(* CODESYS project demo_RECOVERED_2026-10-14T16-49-24.project
   Author: Schneider
   Version: 1.0.0.0

Project tree, tasks and I/O mapping:
  MyController : TM310MM35ECT16U, Schneider Electric, order no. Schneider M310M Target, version 2.0.0.43
    application Application
      libraries: Util, 3.5.19.0 (System); Standard, 3.5.18.0 (System); MC_Basic, 1.10.1.65 (Schneider Electric SA); M310M PLCSystem, * (Schneider Electric)
      task MAST (cyclic, interval T#20ms, priority 15) calls PLC_PRG
      task CommunicationTask (cyclic, interval t#20ms, priority 16) calls nothing
      task MotionTask (cyclic, interval T#4ms, priority 0) calls Motion_PRG, Hidden_PRG
      ImplicitChecks/
        function CheckDivDInt [ST]
        function CheckBounds [ST]
        function CheckLRangeUnsigned [ST]
        function CheckRangeUnsigned [ST]
        function CheckDivReal [ST]
        function CheckDivLReal [ST]
        function CheckRangeSigned [ST]
        function CheckPointer [ST]
        function CheckLRangeSigned [ST]
        function CheckDivLInt [ST]
      program PLC_PRG [ST]
      program Hidden_PRG [ST]
      global variables GVL
      program Motion_PRG [ST]
    Encoders : Encoders, Schneider Electric, version 2.0.0.43
    Cartridge_1 : Cartridge, Schneider Electric, version 2.0.0.43
    IO_Bus : IO bus - TM3, Schneider Electric, version 2.0.0.43
      Module_1 : TM3DI16/G, Schneider Electric, order no. TM3DI16/G, version 1.0.2.2
          input  iwModule_4_IW0 : WORD  // IW0
      Module_2 : TM3DQ16R/G, Schneider Electric, order no. TM3DQ16R/G, version 1.0.2.2
          unmapped channels: QW0
      Module_3 : TM3AI4/G, Schneider Electric, order no. TM3AI4/G, version 1.0.2.2
          settings: KPI Configuration.KPI Configuration = 35; KPI Configuration.KPI Configuration = 160; KPI Configuration.KPI Configuration = 15; KPI Configuration.KPI Configuration = 32; KPI Configuration.KPI Configuration = 78
          input  Application.Motion_PRG.WaterLevel AT %IW3 : INT  // IW0
          input  ibModule_1_IBStatusIW0 : BYTE  // IBStatusIW0
          input  ibModule_1_IBStatusIW1 : BYTE  // IBStatusIW1
          input  ibModule_1_IBStatusIW2 : BYTE  // IBStatusIW2
          input  ibModule_1_IBStatusIW3 : BYTE  // IBStatusIW3
          unmapped channels: %IW4 IW1, %IW5 IW2, IW3
      Module_4 : TM3AQ2/G, Schneider Electric, order no. TM3AQ2/G, version 1.0.2.2
          settings: KPI Configuration.KPI Configuration = 19; KPI Configuration.KPI Configuration = 160; KPI Configuration.KPI Configuration = 15; KPI Configuration.KPI Configuration = 32; KPI Configuration.KPI Configuration = 78
          output qiModule_2_QW1 : INT  // QW1
          input  ibModule_2_IBStatusQW0 : BYTE  // IBStatusQW0
          input  ibModule_2_IBStatusQW1 : BYTE  // IBStatusQW1
          unmapped channels: %QW3 QW0
    EtherCAT_Master_SE : EtherCAT Master SE, Schneider Electric SA, version 4.9.0.3
    Cartridge_2 : Cartridge, Schneider Electric, version 2.0.0.43
    Ethernet_1 : Ethernet Network, Schneider Electric, version 4.3.0.6
        settings: IPAddress = [192,168,0,122]; SubnetMask = [255,255,255,0]; GatewayAddress = [192,168,0,1]; MACAddress = [16#00,16#00,16#00,16#00,16#00,16#00]; IPAddress = [192,168,0,2]; SubnetMask = [255,255,255,0]; GatewayAddress = [0,0,0,0]
      ModbusTCP_Server_Device : ModbusTCP Server Device, Schneider Electric SA, version 4.5.0.1
          input  iwModbusTCP_Server_Device_0 : WORD  // 保持寄存器.保持寄存器
          input  iwModbusTCP_Server_Device_1 : WORD  // 保持寄存器.保持寄存器
          input  iwModbusTCP_Server_Device_2 : WORD  // 保持寄存器.保持寄存器
          input  iwModbusTCP_Server_Device_3 : WORD  // 保持寄存器.保持寄存器
          input  iwModbusTCP_Server_Device_4 : WORD  // 保持寄存器.保持寄存器
          input  iwModbusTCP_Server_Device_5 : WORD  // 保持寄存器.保持寄存器
          input  iwModbusTCP_Server_Device_6 : WORD  // 保持寄存器.保持寄存器
          input  iwModbusTCP_Server_Device_7 : WORD  // 保持寄存器.保持寄存器
          input  iwModbusTCP_Server_Device_8 : WORD  // 保持寄存器.保持寄存器
          input  iwModbusTCP_Server_Device_9 : WORD  // 保持寄存器.保持寄存器
          input  iwModbusTCP_Server_Device_10 : WORD  // 保持寄存器.保持寄存器
          input  iwModbusTCP_Server_Device_11 : WORD  // 保持寄存器.保持寄存器
          input  iwModbusTCP_Server_Device_12 : WORD  // 保持寄存器.保持寄存器
          input  iwModbusTCP_Server_Device_13 : WORD  // 保持寄存器.保持寄存器
          input  iwModbusTCP_Server_Device_14 : WORD  // 保持寄存器.保持寄存器
          input  iwModbusTCP_Server_Device_15 : WORD  // 保持寄存器.保持寄存器
          output qwModbusTCP_Server_Device_0 : WORD  // 输入寄存器.输入寄存器
          output qwModbusTCP_Server_Device_1 : WORD  // 输入寄存器.输入寄存器
          output qwModbusTCP_Server_Device_2 : WORD  // 输入寄存器.输入寄存器
          output qwModbusTCP_Server_Device_3 : WORD  // 输入寄存器.输入寄存器
          output qwModbusTCP_Server_Device_4 : WORD  // 输入寄存器.输入寄存器
          output qwModbusTCP_Server_Device_5 : WORD  // 输入寄存器.输入寄存器
          output qwModbusTCP_Server_Device_6 : WORD  // 输入寄存器.输入寄存器
          output qwModbusTCP_Server_Device_7 : WORD  // 输入寄存器.输入寄存器
          output qwModbusTCP_Server_Device_8 : WORD  // 输入寄存器.输入寄存器
          output qwModbusTCP_Server_Device_9 : WORD  // 输入寄存器.输入寄存器
          output qwModbusTCP_Server_Device_10 : WORD  // 输入寄存器.输入寄存器
          output qwModbusTCP_Server_Device_11 : WORD  // 输入寄存器.输入寄存器
          output qwModbusTCP_Server_Device_12 : WORD  // 输入寄存器.输入寄存器
          output qwModbusTCP_Server_Device_13 : WORD  // 输入寄存器.输入寄存器
          output qwModbusTCP_Server_Device_14 : WORD  // 输入寄存器.输入寄存器
          output qwModbusTCP_Server_Device_15 : WORD  // 输入寄存器.输入寄存器
          unmapped channels: 保持寄存器, 输入寄存器
    Pulse_Generators : Pulse Generators, Schneider Electric, version 2.0.0.43
    Virtual Axis Pool
    COM_1 : Serial COM, Schneider Electric, version 2.0.0.43
    DI : Digital Inputs, Schneider Electric, version 2.0.0.43
        input  iwDI_IW0 : WORD  // IW0
        input  ibDI_IB1 : BYTE  // IB1
    Counters : Counters, Schneider Electric, version 2.0.0.43
    DQ : Digital Outputs, Schneider Electric, version 2.0.0.43
        output qwDQ_QW0 : WORD  // QW0
        output qbDQ_QB1 : BYTE  // QB1
*)

// MyController/Application/GVL
{attribute 'qualified_only'}
VAR_GLOBAL
	rTargetLevel AT %MW0   : REAL := 40.0;    (* 目标水位 %, 占 MW0-1 *)
    rManualValve AT %MW2   : REAL := 0.0;     (* 手动阀开度 %, 占 MW2-3 *)

    (* ===== 状态/报警 (只读供 HMI) ===== *)
	rLevel       AT %MW4   : REAL;     (* 实测水位 %, 占 MW4-5 *)
	rValveCmd    AT %MW6   : REAL;     (* 阀指令 %, 占 MW6-7 *)
END_VAR

// MyController/Application/PLC_PRG
PROGRAM PLC_PRG
VAR
	    (* ===== 周期 ===== *)
    tCycle : TIME := T#100MS;
    rDt    : REAL;                       (* 采样周期, 秒 *)

    (* ===== 物理IO (地址须与 Device IO Mapping 核对) ===== *)
    iLevelRaw AT %IW3    : INT;          (* 水位 4-20mA, 4000..20000 = 0..100% *)
    iValveOut  AT %QW3   : INT;          (* 抽水阀开度 4-20mA, 4000..20000 = 0..100% *)
    bPump      AT %QX4.0 : BOOL;         (* 抽水泵继电器, ON=抽水 *)

    (* ===== HMI / Modbus 设定 (地址可按需调整) ===== *)
    //rTargetLevel AT %MW0   : REAL := 40.0;    (* 目标水位 %, 占 MW0-1 *)
    bAuto        AT %MX102.0 : BOOL := TRUE;    (* 1=自动 0=手动 *)
   // rManualValve AT %MW2   : REAL := 0.0;     (* 手动阀开度 %, 占 MW2-3 *)
    bManualPump  AT %MX106.0 : BOOL := FALSE;   (* 手动泵 ON *)

    (* ===== 状态/报警 (只读供 HMI) ===== *)
	//rLevel       AT %MW4   : REAL;     (* 实测水位 %, 占 MW4-5 *)
	//rValveCmd    AT %MW6   : REAL;     (* 阀指令 %, 占 MW6-7 *)
    bPumpCmd     AT %MX114.0 : BOOL;     (* 泵指令 *)
    bSensorFault AT %MX114.1 : BOOL;     (* 传感器故障 *)
    bAlarm       AT %MX114.2 : BOOL;     (* 总报警 *)

    (* ===== 量程 (INT) ===== *)
    iRawMin : INT := 4000;
    iRawMax : INT := 20000;

    (* ===== PID 内部 ===== *)
    rError, rPrevError, rInt, rDeriv, rPD, rOut : REAL;

    (* ===== PID 参数 (待整定, 见文档) ===== *)
    //rKp : REAL := 3.0;
   // rKi : REAL := 0.1;     (* 1/s, 抵消自然入流静差; 积分对象 Ki 勿过大 *)
   // rKd : REAL := 0.0;
	rKp AT %MW20 : REAL := 3.0;      (* 占 MW20-21, 默认值(上电/未使能时用) *)
    rKi AT %MW22 : REAL := 0.5;      (* 占 MW22-23 *)
    rKd AT %MW24 : REAL := 0.0;      (* 占 MW24-25 *)
    bPidTune : BOOL := FALSE;        (* 1=采用 Modbus 传入的 Kp/Ki/Kd, 0=用上面默认 *)

    (* ===== 联锁阈值 (%, 工程量) ===== *)
    rLvlHH      : REAL := 95.0;   (* 高高: 最大抽水降压 *)
    rLvlLL      : REAL := 5.0;    (* 低低: 停泵防干抽, 靠自流回涨 *)
    rPumpOnThr  : REAL := 3.0;    (* 阀开度>3% 开泵 *)
    rPumpOffThr : REAL := 1.0;    (* 阀开度<1% 关泵(防憋压) *)
	
END_VAR

rDt := TIME_TO_REAL(tCycle) / 1000;   (* 0.1 s *)
(* ===== Modbus 读入: 上位机 -> PLC 设定值 ===== *)
(* REAL 占 2 字, 低字在前(Device_0=低字, 与现有 rLevel 映射顺序一致) *)
%MW0 := iwModbusTCP_Server_Device_0;   (* rTargetLevel 低字 *)
%MW1 := iwModbusTCP_Server_Device_1;   (* rTargetLevel 高字 *)
%MW2 := iwModbusTCP_Server_Device_6;   (* rManualValve 低字 (可选) *)
%MW3 := iwModbusTCP_Server_Device_7;   (* rManualValve 高字 (可选) *)
bAuto       := iwModbusTCP_Server_Device_10.0;   (* 提取 bit0 *)
bManualPump := iwModbusTCP_Server_Device_10.1;   (* 提取 bit1 *)
bPidTune    := iwModbusTCP_Server_Device_10.2;   (* 提取 bit2 *)

(* 仅当使能位置 1 时, 才用 Modbus 传入的 PID 参数覆盖默认值 *)
IF bPidTune THEN
    %MW20 := iwModbusTCP_Server_Device_2;    (* rKp 低字 *)
    %MW21 := iwModbusTCP_Server_Device_3;    (* rKp 高字 *)
    %MW22 := iwModbusTCP_Server_Device_4;    (* rKi 低字 *)
    %MW23 := iwModbusTCP_Server_Device_5;    (* rKi 高字 *)
    %MW24 := iwModbusTCP_Server_Device_12;   (* rKd 低字 *)
    %MW25 := iwModbusTCP_Server_Device_13;   (* rKd 高字 *)

    (* 安全钳制: 防止写入过大值导致剧烈振荡 *)
    rKp := LIMIT(0.0, rKp, 20.0);
    rKi := LIMIT(0.0, rKi, 5.0);
    rKd := LIMIT(0.0, rKd, 10.0);
END_IF
(* bPidTune=0 时不覆盖, rKp/rKi/rKd 保持声明里的默认(或上一次使能写入的值) *)

(* ---------- 1. 传感器自检 + 水位标定 ---------- *)
IF (iLevelRaw < iRawMin - 200) OR (iLevelRaw > iRawMax + 200) THEN
    bSensorFault := TRUE;
ELSE
    bSensorFault := FALSE;
END_IF
GVL.rLevel := LIMIT(0.0,
    (INT_TO_REAL(iLevelRaw - iRawMin) / 16000.0) * 100.0, 100.0);

(* ---------- 2. 联锁 (最高优先级) ---------- *)
IF bSensorFault THEN
    (* 传感器故障: 停泵关阀+报警 (自然入流会缓慢上升, 需人工干预) *)
    bPumpCmd  := FALSE;
    GVL.rValveCmd := 0.0;
    rInt      := 0.0;
ELSIF (GVL.rLevel >= rLvlHH) THEN
    (* 高高液位: 最大抽水快速降压 *) 
    bPumpCmd  := TRUE;
    GVL.rValveCmd := 100.0;
    rInt      := 0.0;
ELSIF (GVL.rLevel <= rLvlLL) THEN
    (* 低低液位: 停抽防干抽, 靠自然入流回涨 *)
    bPumpCmd  := FALSE;
    GVL.rValveCmd := 0.0;
    rInt      := 0.0;
ELSE
    (* ---------- 3. PID (阀在抽水侧: 偏高->开阀抽水) ---------- *)
    rError := GVL.rLevel - GVL.rTargetLevel;            (* PV - SP, 正=偏高需抽水 *)
    rDeriv := (rError - rPrevError) / rDt;
    rPD    := rKp * rError + rKd * rDeriv;
    rOut   := rPD + rKi * rInt;

    (* 抗积分饱和: 输出饱和且误差同向时冻结积分 *)
    IF NOT ((rOut > 100.0 AND rError > 0.0) OR (rOut < 0.0 AND rError < 0.0)) THEN
        rInt := rInt + rError * rDt;
        rInt := LIMIT(-100.0, rInt, 100.0);
    END_IF
    GVL.rValveCmd := LIMIT(0.0, rPD + rKi * rInt, 100.0);
    rPrevError := rError;

    (* ---------- 4. 泵启停迟滞 (保护继电器+防憋压) ---------- *)
    IF bPumpCmd THEN
        IF GVL.rValveCmd < rPumpOffThr THEN bPumpCmd := FALSE; END_IF
    ELSE
        IF GVL.rValveCmd > rPumpOnThr  THEN bPumpCmd := TRUE;  END_IF
    END_IF
END_IF

(* ---------- 5. 手动模式 (含无扰切换: 积分跟踪手动阀开度) ---------- *)
IF NOT bAuto THEN
    GVL.rValveCmd := LIMIT(0.0, GVL.rManualValve, 100.0);
    bPumpCmd  := bManualPump;
    IF rKi <> 0.0 THEN
        rInt := (GVL.rValveCmd - rKp * (GVL.rLevel - GVL.rTargetLevel)) / rKi;
        rInt := LIMIT(-100.0, rInt, 100.0);
    END_IF
    rPrevError := GVL.rLevel - GVL.rTargetLevel;
END_IF

(* ---------- 6. 输出标定与写入 ---------- *)
iValveOut := LIMIT(iRawMin,
    iRawMin + REAL_TO_INT(GVL.rValveCmd / 100.0 * 16000.0), iRawMax);
bPump := bPumpCmd AND NOT bSensorFault;

(* ---------- 7. 报警汇总 ---------- *)
bAlarm := bSensorFault OR (GVL.rLevel >= rLvlHH) OR (GVL.rLevel <= rLvlLL);

(* ===== Modbus 写出: PLC -> 上位机 只读状态 ===== *)
qwModbusTCP_Server_Device_2 := %MW4;   (* rLevel 低字 *)
qwModbusTCP_Server_Device_3 := %MW5;   (* rLevel 高字 *)
qwModbusTCP_Server_Device_4 := %MW6;   (* rValveCmd 低字 *)
qwModbusTCP_Server_Device_5 := %MW7;   (* rValveCmd 高字 *)
(* bit0=bAuto, bit1=bPumpCmd, bit2=bSensorFault, bit3=bAlarm, bit4=bPump *)
(* 直接给 WORD 的指定位赋值，0 警告，执行效率极高 *)
qwModbusTCP_Server_Device_8.0 := bAuto;         (* 第 0 位赋值 *)
qwModbusTCP_Server_Device_8.1 := bPumpCmd;      (* 第 1 位赋值 *)
qwModbusTCP_Server_Device_8.2 := bSensorFault;  (* 第 2 位赋值 *)
qwModbusTCP_Server_Device_8.3 := bAlarm;        (* 第 3 位赋值 *)
qwModbusTCP_Server_Device_8.4 := bPump;         (* 第 4 位赋值 *)
qwModbusTCP_Server_Device_10 := %MW20;   (* rKp 低字 *)
qwModbusTCP_Server_Device_11 := %MW21;   (* rKp 高字 *)
qwModbusTCP_Server_Device_12 := %MW22;   (* rKi 低字 *)
qwModbusTCP_Server_Device_13 := %MW23;   (* rKi 高字 *)
qwModbusTCP_Server_Device_14 := %MW24;   (* rKd 低字 *)
qwModbusTCP_Server_Device_15 := %MW25;   (* rKd 高字 *)

END_PROGRAM

// MyController/Application/Motion_PRG
PROGRAM Motion_PRG
VAR
	WaterLevel : INT := 0;
	Threshold : INT := 0;
	testval : INT := 0;
	switchon : word:=0;
END_VAR

WaterLevel := WaterLevel;
//Threshold := testval;

END_PROGRAM

// MyController/Application/Hidden_PRG
PROGRAM Hidden_PRG
VAR
   bStartRunFlag:BOOL:=FALSE;
END_VAR

MC_IN_MotionCalculate();

END_PROGRAM

// MyController/Application/ImplicitChecks/CheckDivDInt
// 隐式生成代码:不需要编辑
FUNCTION CheckDivDInt : DINT
VAR_INPUT
	divisor:DINT;
END_VAR

// 隐式生成代码:只是实现代码的建议
IF divisor = 0 THEN
	CheckDivDInt:=1;
ELSE
	CheckDivDInt:=divisor;
END_IF;

END_FUNCTION

// MyController/Application/ImplicitChecks/CheckBounds
// 隐式生成代码:不需要编辑
FUNCTION CheckBounds : DINT
VAR_INPUT
	index, lower, upper: DINT;
END_VAR

// 隐式生成代码:只是实现代码的建议
IF  index < lower THEN
	CheckBounds := lower;
ELSIF  index > upper THEN
	CheckBounds := upper;
ELSE  
	CheckBounds := index;
END_IF

(*还可以设置断点,日志信息或其他.比如在异常处停止:
Add CmpApp.library, SysExcept.library and SysTypes2_Itf as newest.
Declaration:
VAR
    _pApp : POINTER TO CmpApp.APPLICATION;
    _result   : SysTypes.RTS_IEC_RESULT;
END_VAR

Implementation:
_pApp := AppGetCurrent(pResult:=_result);
IF  index < lower THEN
        CheckBounds := lower;
        IF _pApp <> 0 THEN
                AppGenerateException(pApp:=_pApp, ulException:=RtsExceptions.RTSEXCPT_ARRAYBOUNDS);
        END_IF
ELSIF  index > upper THEN
        CheckBounds := upper;
        IF _pApp <> 0 THEN
                AppGenerateException(pApp:=_pApp,   ulException:=RtsExceptions.RTSEXCPT_ARRAYBOUNDS);
        END_IF
ELSE  
        CheckBounds := index;
END_IF
*)

END_FUNCTION

// MyController/Application/ImplicitChecks/CheckLRangeUnsigned
// 隐式生成代码:不需要编辑
FUNCTION CheckLRangeUnsigned : ULINT
VAR_INPUT
	value, lower, upper: ULINT;
END_VAR

// 隐式生成代码:只是实现代码的建议
IF (value < lower) THEN
	CheckLRangeUnsigned := lower;
ELSIF(value > upper) THEN
	CheckLRangeUnsigned := upper;
ELSE
	CheckLRangeUnsigned := value;
END_IF

END_FUNCTION

// MyController/Application/ImplicitChecks/CheckRangeUnsigned
// 隐式生成代码:不需要编辑
FUNCTION CheckRangeUnsigned : UDINT
VAR_INPUT
	value, lower, upper: UDINT;
END_VAR

// 隐式生成代码:只是实现代码的建议
IF (value < lower) THEN
	CheckRangeUnsigned := lower;
ELSIF(value > upper) THEN
	CheckRangeUnsigned := upper;
ELSE
	CheckRangeUnsigned := value;
END_IF

END_FUNCTION

// MyController/Application/ImplicitChecks/CheckDivReal
// 隐式生成代码:不需要编辑
FUNCTION CheckDivReal : REAL
VAR_INPUT
	divisor:REAL;
END_VAR

// 隐式生成代码:只是实现代码的建议
IF divisor = 0 THEN
	CheckDivReal:=1;
ELSE
	CheckDivReal:=divisor;
END_IF;

END_FUNCTION

// MyController/Application/ImplicitChecks/CheckDivLReal
// 隐式生成代码:不需要编辑
FUNCTION CheckDivLReal : LREAL
VAR_INPUT
	divisor:LREAL;
END_VAR

// 隐式生成代码:只是实现代码的建议
IF divisor = 0 THEN
	CheckDivLReal:=1;
ELSE
	CheckDivLReal:=divisor;
END_IF;

END_FUNCTION

// MyController/Application/ImplicitChecks/CheckRangeSigned
// 隐式生成代码:不需要编辑
FUNCTION CheckRangeSigned : DINT
VAR_INPUT
	value, lower, upper: DINT;
END_VAR

// 隐式生成代码:只是实现代码的建议
IF (value < lower) THEN
	CheckRangeSigned := lower;
ELSIF(value > upper) THEN
	CheckRangeSigned := upper;
ELSE
	CheckRangeSigned := value;
END_IF

END_FUNCTION

// MyController/Application/ImplicitChecks/CheckPointer
// 隐式生成代码:不需要编辑
FUNCTION CheckPointer : POINTER TO BYTE
VAR_INPUT 
	ptToTest : POINTER TO BYTE; // 指针的目标地址
	iSize : DINT;		        // 指针指向的类型大小.(例如:POINTER TO ARRAY [0..9] OF INT为20)
	iGran : DINT;		        // 指针访问的粒度,即指针指向的类型中最大的非结构数据类型的大小.(例如: POINTER TO ARRAY [0..9] OF INT为2)
	bWrite: BOOL;		        // 标识读或写权限.TRUE = 写权限.
END_VAR

// 没有标准的实现方式.在此处输入代码
CheckPointer := ptToTest;

END_FUNCTION

// MyController/Application/ImplicitChecks/CheckLRangeSigned
// 隐式生成代码:不需要编辑
FUNCTION CheckLRangeSigned : LINT
VAR_INPUT
	value, lower, upper: LINT;
END_VAR

// 隐式生成代码:只是实现代码的建议
IF (value < lower) THEN
	CheckLRangeSigned := lower;
ELSIF(value > upper) THEN
	CheckLRangeSigned := upper;
ELSE
	CheckLRangeSigned := value;
END_IF

END_FUNCTION

// MyController/Application/ImplicitChecks/CheckDivLInt
// 隐式生成代码:不需要编辑
FUNCTION CheckDivLInt : LINT
VAR_INPUT
	divisor:LINT;
END_VAR

// 隐式生成代码:只是实现代码的建议
IF divisor = 0 THEN
	CheckDivLInt:=1;
ELSE
	CheckDivLInt:=divisor;
END_IF;

END_FUNCTION
